// TIA Portal V21 export
FUNCTION "FC_AnaCaseReal" : Int   // FC14, SCL
TITLE = Analyzer: CASE without ELSE, REAL compared with =
{ S7_Optimized_Access := 'TRUE' }
// Rule C26i: the CASE has no ELSE, and a REAL is compared with =
// stored: SetENOAutomatically false
   VAR_INPUT
      Mode : Int;   // Mode
      Level : Real;   // Level
   END_VAR
   VAR_TEMP
      Code : Int;   // Result code
   END_VAR
BEGIN

       #Code := 0;
       CASE #Mode OF
           1:
               #Code := 10;
           2:
               #Code := 20;
       END_CASE;
       IF #Level = 1.5 THEN
           #Code := #Code + 1;
       END_IF;
       #FC_AnaCaseReal := #Code;
END_FUNCTION
